{attribute 'qualified_only'}
{attribute 'strict'}
TYPE E_FaultCode :
(
	FC_NONE,
	FC_EMERGENCY_STOP,
	FC_EXIT_TIMEOUT
);
END_TYPE

(* stored: Version 1.1.0.1, ProductVersion 3.1.4024.16
   DUT E_FaultCode: Id {96265e21-0ab7-464f-9ca5-fa08e81b9f3a} *)
